(* IEC 61131-3 sources: axsharp/src/ix.examples/hello.world.console/hello.world.console.plc/src, 2 files *)

(* ---- configuration.st ---- *)
CONFIGURATION MyConfiguration
    TASK Main(Interval := T#1000ms, Priority := 1);
    PROGRAM P1 WITH Main: MyProgram;

    VAR_GLOBAL
        Counter : ULINT;
        HelloWorld : STRING := 'Hello world';
    END_VAR
END_CONFIGURATION

(* ---- program.st ---- *)
PROGRAM MyProgram
    VAR_EXTERNAL
        Counter : ULINT;
        HelloWorld : STRING;
    END_VAR

    Counter := Counter + ULINT#1;
    IF(HelloWorld = 'RESET-COUNTER') THEN
        Counter := ULINT#0;
    END_IF;
END_PROGRAM
